TYPE ST_Node :
STRUCT
	/// Axis ID 
	nAxisId: DWORD;
	pMover: POINTER TO ST_Axis := null;
	pPremover: POINTER TO ST_Axis := null;
	pAftermover: POINTER TO ST_Axis := null;
END_STRUCT
END_TYPE

(* stored: Version 1.1.0.1, ProductVersion 3.1.4024.12
   DUT ST_Node: Id {80eb2b5e-3aae-4806-b66a-875c102b1961} *)
